INTERFACE I_Safety

PROPERTY PUBLIC doorLock : BOOL
GET
END_GET
SET
END_SET
END_PROPERTY

PROPERTY inHold : BOOL
GET
END_GET
END_PROPERTY

PROPERTY isDoorSafe : BOOL
GET
END_GET
END_PROPERTY

PROPERTY isDoorUsed : BOOL
GET
END_GET
END_PROPERTY

PROPERTY isSafe : BOOL
GET
END_GET
END_PROPERTY

END_INTERFACE

(* stored: Version 1.1.0.1, ProductVersion 3.1.4024.12
   Itf I_Safety: Id {baf468b0-bf3f-48fa-95b7-6b03bb61a91e}
   Property doorLock: Id {d4e5cdd7-10d8-44cf-bb45-8aa3265e1026}
   Get Get: Id {5c76633d-644a-496d-b5cd-abdc98f6241e}
   Set Set: Id {1b9dece8-2d3a-4d2f-8de3-3e0b3ae99ccb}
   Property inHold: Id {f8a6d36b-536e-44e4-baaf-e25567ad39bb}
   Get Get: Id {219ec9ae-a0d8-48ab-a07b-fffffa96e448}
   Property isDoorSafe: Id {7de6b713-a2a8-42a8-bfcb-32f6ff9b2c2d}
   Get Get: Id {bd00fb9e-51bb-45e4-8cef-d833d52344b3}
   Property isDoorUsed: Id {09b63899-f848-45a5-a99a-c9dc8840c4aa}
   Get Get: Id {2b8cc24d-caf8-4e66-9172-d009411c7ef4}
   Property isSafe: Id {6bbdf64d-2bcf-46ff-b423-deaa4449811c}
   Get Get: Id {036d2111-6b1d-40c8-9041-e6c712f75f61} *)
